       #instGetIoPart(ID := #hwID,   //read data from process image
                      OFFSET := #portAddr,
                      LEN := #statIOsize,
                      STATUS => #statIoPartStatus,
                      ERROR => #statIoPartError,
                      INPUTS := #statAnt);
       #statAntStatus := #statAnt[#INDEX_ANT_STATUS];    //status byte
       #statPresence := #statAntStatus.%X5;    //Presence bit. Transponder on field
   END_REGION

   REGION Check antenna status
       IF #statAnt[#INDEX_RFID_ERROR] <> 0 AND #statBusy THEN
           #tempStatus.%W0 := BYTE_TO_WORD(#statAnt[#INDEX_RFID_ERROR]);    //error_BLK
           #tempStatus.%W1 := #STATUS_ERROR_IDENT_RFID;                    //identifier rfid errors
           #statBusy := false;
           #tempDone := false;
           #tempError := TRUE;
           #statState := #STATE_IDLE;
       END_IF;
   END_REGION

   REGION Check execute
       REGION Idle
           IF NOT #execute THEN
               #tempDone := false;
               #tempError := false;
               #tempStatus := 0;
           END_IF;
       END_REGION

       REGION Job executed
           IF #execute AND #execute <> #statExecuteReq THEN //Positive Edge for antenna on
               #statBusy := TRUE;                              //Block active
               #tempDone := FALSE;                             //reset all output parameters
               #tempError := FALSE;
               #tempStatus := #STATUS_NO_JOB;
               IF #antennaState THEN                          //if antenna then activate the ANTENNA_ON process
                   #statState := #STATE_ANTENNA_ON;
               ELSIF NOT #antennaState THEN                   //if not antenna then activate the ANTENNA_OFF process 
                   #statState := #STATE_ANTENNA_OFF;
               END_IF;

           END_IF;
       END_REGION
       #statExecuteReq := #execute;
   END_REGION

   REGION State machine
       CASE #statState OF
           #STATE_IDLE:
               ;

           #STATE_ANTENNA_ON:  //Antenna_on
               //Antenna on process
               #statAntStatus.%X4 := false;                        //Reset Byte 0, bit 4
               #statSent[#INDEX_SEND_CMD] := #CMD_ANTENNA_ON;
               #instSetIoPart(ID := #hwID,                         //Write data into process image
                              OFFSET := #portAddr,
                              LEN := #statIOsize,
                              STATUS => #statIoPartStatus,
                              ERROR => #statIoPartError,
                              OUTPUTS := #statSent);
               IF NOT #statIoPartError AND #statAnt[#INDEX_RFID_ERROR] = 0 THEN
                   #statState := #STATE_READY;
               ELSIF #statIoPartError THEN
                   #tempError := true;
                   #statBusy := FALSE;
                   #tempStatus.%W0 := DWORD_TO_WORD(#statIoPartStatus);//error_BLK
                   #tempStatus.%W1 := #STATUS_ERROR_IDENT_BLOCK;                    //identifier block errors
                   #statState := #STATE_IDLE;
               END_IF;

           #STATE_ANTENNA_OFF:
               //Antenna off process
               #statAntStatus.%X4 := true;                         //set Byte 0, bit 4
               #statSent[#INDEX_SEND_CMD] := #CMD_ANTENNA_OFF;
               #instSetIoPart(ID := #hwID,                         //Write data into process image
                              OFFSET := #portAddr,
                              LEN := #statIOsize,
                              STATUS => #statIoPartStatus,
                              ERROR => #statIoPartError,
                              OUTPUTS := #statSent);
               IF NOT #statIoPartError AND #statAnt[#INDEX_RFID_ERROR] = 0 THEN
                   IF #statAntStatus = #CMD_ANTENNA_OFF THEN    //if status_byte=16#10 then antenna off
                       #statState := #STATE_READY;
                   END_IF;
               ELSIF #statIoPartError THEN
                   #tempError := true;
                   #statBusy := FALSE;
                   #tempStatus.%W0 := DWORD_TO_WORD(#statIoPartStatus);    //error_BLK
                   #tempStatus.%W1 := #STATUS_ERROR_IDENT_BLOCK;   //identifier block errors
                   #statState := #STATE_IDLE;
               END_IF;

           #STATE_READY:
               #tempDone := true;
               #statBusy := FALSE;
               #statState := #STATE_IDLE;
           ELSE
               #statState := #STATE_IDLE;
       END_CASE;
   END_REGION

   REGION Update output interface 
       #done := #tempDone;
       #busy := #statBusy;
       #error := #tempError;
       #status := #tempStatus;
       #presence := #statPresence;
   END_REGION
END_FUNCTION_BLOCK

FUNCTION_BLOCK "LIOLink_RF200_WriteTag"   // FB6, SCL
TITLE = LIOLink_RF200_WriteTag
{ S7_Optimized_Access := 'TRUE' }
AUTHOR : SIOS
FAMILY : LIOLink
VERSION : 2.4
// Writes tags on SIMATIC RF200 readers via IO-Link
   VAR_INPUT
      execute : Bool;   // Execute function
      addrTag : Word;   // Start address of data on tag
      length : Word;   // Length of data to be written
      hwID : HW_SUBMODULE;   // Hardware identifier of IO-Link communication module
      portAddr : Int;   // Start address of port
      "version" : USInt := 11;   // IO-Link version of the reader; 11: IO-Link V1.1, 10: IO-Link V1.0
   END_VAR
   VAR_OUTPUT
      done : Bool;   // TRUE: job done
      busy : Bool;   // FALSE: no job, TRUE: job in progress
      error : Bool;   // FALSE: no error, TRUE: error
      status : DWord;   // Error Status
      presence : Bool;   // Tag on antenna field
   END_VAR
   VAR_IN_OUT
      identData : Variant;   // Data to write in
   END_VAR
   VAR
      instTonR : TONR_TIME;   // Tag has left antenna field detection timer
      statState : Int;   // Main State Machine Index
      statTimerIn : Bool;   // Tag has left antenna field detection timer - Start Tag
      statTimerR : Bool;   // Tag has left antenna field detection timer - Reset Tag
      statTimerPt : Time := T#5S;   // Tag has left antenna field detection timer - Detection time
      statStatusByte : Byte;   // First received Byte from process image
      statDat : Array[0..#UPPER_BOUND_IO_FIELD] of Byte;   // Sent data
      statRecDat : Array[0..#UPPER_BOUND_IO_FIELD] of Byte;   // Received data
      statPresence : Bool;   // TRUE: Transponder on field
      statExecuteReq : Bool;   // State of execute input of last cycle
      statLength : DInt;   // Length of read Data
      statAddr : Word;   // Address of Tag
      statWriteOffset : Int;   // Data offset for write function
      statPresenceFf : Bool;   // Transpnder status of last cycle
      statWriteData : Array[0..#UPPER_BOUND_MAX_DATA_FIELD] of Byte;   // Data to write to tag
      statDiffToIOsizeNetto : Int;   // Difference to full IO size
      statBytemove : Int;   // Shift value for data
      statDone : Bool;   // TRUE: job done
      statBusy : Bool;   // FALSE: no job, TRUE: job in progress
      statError : Bool;   // FALSE: no error, TRUE: error
      instSetIoPart : SETIO_PART;   // Instance for PIQ writing
      statIoPartError : Bool;   // TRUE: data in process image is invalid
      statIoPartStatus : DWord;   // Status for IO access
      instGetIoPart : GETIO_PART;   // Instance for PII reading
      statReturnMoveBlkVar : Int;   // Return Value of Block Move
      statIOsize : USInt;   // Size of the IO-Link Master PII
      statIOsizeNetto : USInt;   // Size of the IO-Link Master PAE without header
   END_VAR
   VAR_TEMP
      tempStatus : DWord;   // Auxiliary tag for status output
   END_VAR
   VAR CONSTANT
      IOL_V10 : USInt := 10;   // Identifier IO-Link version 1.0
      IOL_V11 : USInt := 11;   // Identifier IO-Link version 1.1
      LEN_DATA_V10 : USInt := 8;   // Length of user data for IO-Link version 1.0
      LEN_DATA_V11 : USInt := 32;   // Length of user data for IO-Link version 1.1
      UPPER_BOUND_IO_FIELD : USInt := 31;   // Upper bound of Input and Output fields
      UPPER_BOUND_MAX_DATA_FIELD : UInt := 1999;   // Upper bound of the data field of a RFID Tag
      DATA_HEADER_SIZE : USInt := 4;   // IO-Link Header Size for version 1.0 and 1.1
      STATUS_ERROR_IDENT_BLOCK : Word := 16#0001;   // Error Identification for block internal faults
      STATUS_ERROR_IDENT_RFID : Word := 16#0011;   // Error Identification for RFID reader faults
      STATUS_NO_JOB : Word := 16#0000;   // No job requested
      STATUS_ERROR_TAG_HAS_LEFT : Word := 16#8101;   // Error - the RFID tag has left the reader
      STATUS_ERROR_STILL_ACTIVE : Word := 16#8102;   // Error - block still busy, no further request possible
      STATUS_ERROR_LENGTH : Word := 16#8104;   // Error - requested length is less than 0
      STATE_IDLE : Int := 0;   // State Machine - Idle State
      STATE_WRITE : Int := 2;   // State Machine - Read Tag
      STATE_TELEGRAM : Int := 1;   // State Machine - Prepare telegram
      STATE_ERROR : Int := 3;   // State Machine - Error State
      DETECTION_TIME_TAG_OFF_FIELD : Time := T#5S;   // Tag has left antenna field detection time
      CMD_WRITE : Byte := 16#01;   // Command to read data
      CMD_RESET : Byte := 16#00;   // Command to reset
      INDEX_CMD : USInt := 0;   // Index in DataField - Command
      INDEX_RFID_ERROR : USInt := 1;   // Index in DataField - Error
      INDEX_ADDR_HIGH : USInt := 2;   // Index in DataField - Address High Byte
      INDEX_ADDR_LOW : USInt := 3;   // Index in DataField - Address Low Byte
      INDEX_SOURCE_DATA : DInt := 4;   // Index in Data Field - Start of netto Data
      INDEX_REC_STATUS : DInt := 0;   // Index in Received DataField - Status
   END_VAR
   // statRecDat[0] := 16#0000;
   // statRecDat[1] := 16#0000;
   // statRecDat[2] := 16#00FF;
   // statRecDat[3] := 16#00FF;
BEGIN
   REGION BLOCK INFO HEADER
       //===============================================================================
       // Siemens / (c)Copyright 2022
       //-------------------------------------------------------------------------------
       // Title:            LIOLink_RF200_WriteTag
       // Function:         Writes tags on SIMATIC RF200 readers via IO-Link
       // Library:          LIOLink
       // Author:           Siemens Industry Online Support
       // Tested with:      CPU 1513-1 PN FW 2.8
       // Engineering:      TIA Portal V16
       // Restrictions:     --
       // Requirements:     --
       //-------------------------------------------------------------------------------
       // Change log table:
       // Version  | Date       | Expert in charge       | Changes applied
       //----------|------------|------------------------|------------------------------
       // 01.00.00 | 01.03.2015 | Online Support         | First release
       // 01.01.00 | 01.12.2016 | Online Support         | Upgrade to TIA Portal V14
       // 02.00.00 | 01.09.2017 | Online Support         | Upgrade to TIA Portal V14 SP1
       //                                                | Implementation of Programming styleguide
       //                                                | Added support for IO-Link V1.1 readers
       // 02.01.00 | 01.12.2017 | Online Support         | Bug fixes and performance improvements
       // 02.02.00 | 01.03.2020 | Online Support         | Upgrade to TIA Portal V16
       // 02.03.00 | 22.09.2020 | Online Support         | Integrated FB into LIOLink library
       //                                                | Renamed FB to LIOLink_RF200_WriteTag
       //                                                | Combined FBs for IO-Link V1.0 and V1.1
       //                                                | Minor bug fixes
       // 02.04.00 | 04.10.2022 | SUP SPH                | Optimization                                               
       //===============================================================================
   END_REGION

   REGION Check version
       IF #version = #IOL_V11 THEN   //determine IO-Link reader version (1.0/1.1) to set offsets
           #statIOsize := #LEN_DATA_V11;
           #statIOsizeNetto := #LEN_DATA_V11 - #DATA_HEADER_SIZE;
       ELSE
           #statIOsize := #LEN_DATA_V10;
           #statIOsizeNetto := #LEN_DATA_V10 - #DATA_HEADER_SIZE;
       END_IF;
   END_REGION

   REGION Get PII
       //read data from process image
       #instGetIoPart(ID := #hwID,
                      OFFSET := #portAddr,
                      LEN := #statIOsize,
                      STATUS => #statIoPartStatus,
                      ERROR => #statIoPartError,
                      INPUTS := #statRecDat);

       #statStatusByte := #statRecDat[#INDEX_REC_STATUS];    //Status Byte
       #statPresence := #statStatusByte.%X5;   //Presence bit. Transponder on field
   END_REGION

   REGION Check execute
       REGION Idle
           IF NOT #execute THEN
               #statDone := false;
               #statBusy := false;
               #statError := false;
               #tempStatus := #STATUS_NO_JOB;
           END_IF;
       END_REGION

       #statDiffToIOsizeNetto := WORD_TO_INT(#length) MOD #statIOsizeNetto;
       REGION Job requested
           IF #execute AND #execute <> #statExecuteReq THEN    //Positive edge for reading of data
               IF NOT #statBusy THEN
                   #statAddr := #addrTag;    //Transpoder Adress
                   #statLength := WORD_TO_DINT(#length);   //Length of read Data
                   #statState := #STATE_WRITE;
                   #statBusy := TRUE;
                   #statDone := FALSE;   //reset all the output parameters                                   
                   #statError := FALSE;
                   #tempStatus := #STATUS_NO_JOB;
                   #statWriteOffset := 0;
                   #statBytemove := 0;
                   //next step >> send write command
               ELSE
                   #tempStatus.%W0 := #STATUS_ERROR_STILL_ACTIVE;    //block is still active
                   #tempStatus.%W1 := #STATUS_ERROR_IDENT_BLOCK;   //Error identifier for block errors
                   #statState := #STATE_ERROR;
               END_IF;
               IF #length < USINT_TO_WORD(#statIOsizeNetto) THEN
                   #tempStatus.%W0 := #STATUS_ERROR_LENGTH;    //length too short
                   #tempStatus.%W1 := #STATUS_ERROR_IDENT_BLOCK;   //identifier rfid errors
                   #tempStatus := #tempStatus;
                   #statState := #STATE_ERROR;
               END_IF;
           END_IF;
       END_REGION
       #statExecuteReq := #execute;
   END_REGION

   REGION Tag presence detection
       IF NOT #statPresence AND #statPresence <> #statPresenceFf THEN    //the tag has left the antenna  field
           IF NOT #statDone THEN
               #statTimerIn := true;   //wait 5 sec
               #statTimerR := false;
           END_IF;
       END_IF;
       #statPresenceFf := #statPresence;
       IF #statPresence THEN
           #statTimerR := true;
           #statTimerIn := false;
       END_IF;
   END_REGION

   REGION State machine
       CASE #statState OF
           #STATE_IDLE:
               #statWriteOffset := 0;    //offset of puffer must be reseted
               #statBusy := false;
               #statTimerIn := false;

           #STATE_WRITE:
               IF #statLength > 0 THEN
                   #statDat[#INDEX_CMD] := #CMD_WRITE;   //Set write command
                   #statDat[#INDEX_ADDR_HIGH] := #statAddr.%B1;    //Adr-H
                   #statDat[#INDEX_ADDR_LOW] := #statAddr.%B0;   //Adr-L
                   VariantGet(SRC := #identData,
                              DST => #statWriteData);

                   #statReturnMoveBlkVar := MOVE_BLK_VARIANT(SRC := #statWriteData,
                                                             COUNT := #statIOsizeNetto,
                                                             SRC_INDEX := #statWriteOffset - #statBytemove,
                                                             DEST_INDEX := #INDEX_SOURCE_DATA,
                                                             DEST => #statDat);
                   //Just #statIOsizeNetto Bytes are reserved for every transfer
               END_IF;
               IF NOT #statIoPartError THEN
                   #statState := #STATE_TELEGRAM;    //Telegram: Edit the read data
               END_IF;

           #STATE_TELEGRAM:
               IF #statLength > 0 THEN   //Only when length of data>0 can continue  
                   IF #statStatusByte.%X6 THEN   //IF RFID error has occured
                       #tempStatus.%W0 := #statRecDat[#INDEX_RFID_ERROR];
                       #tempStatus.%W1 := #STATUS_ERROR_IDENT_RFID;    //Error identifier for RFID errors
                       #statState := #STATE_ERROR;
                   END_IF;

                   //-------------------------- write command is ready------------------------------------------------//
                   IF #statStatusByte.%X7 AND #statStatusByte.%X0 THEN
                       IF #statRecDat[#INDEX_ADDR_HIGH] = #statAddr.%B1 AND #statRecDat[#INDEX_ADDR_LOW] = #statAddr.%B0 THEN //received ADR must be ==sent ADR

                           IF NOT #statIoPartError THEN
                               IF #statStatusByte.%X7 AND NOT #statStatusByte.%X6 THEN
                                   #statLength := #statLength - #statIOsizeNetto;
                                   IF #statDiffToIOsizeNetto <> 0 AND #statLength < #statIOsizeNetto THEN
                                       #statBytemove := #statIOsizeNetto - #statDiffToIOsizeNetto;
                                   END_IF;
                                   //if len is not dividable with #statIOsizeNetto the adr offset has to be changed that the last (length < #statIOsizeNetto) command is done right
                                   #statWriteOffset := #statWriteOffset + #statIOsizeNetto;                                   //offset must be changed
                                   #statAddr := INT_TO_WORD(WORD_TO_INT(#statAddr) + USINT_TO_INT(#statIOsizeNetto) - #statBytemove);     //Change the ADR on Transponder(#statIOsizeNetto Bytes)       
                                   #statState := #STATE_WRITE;                      //Start a new write command
                               ELSE
                                   #statState := #STATE_IDLE;
                               END_IF;
                           ELSE
                               #tempStatus.%W0 := DWORD_TO_WORD(#statIoPartStatus);    //Error has to BLKMOV occured
                               #tempStatus.%W1 := #STATUS_ERROR_IDENT_BLOCK;   //functions-Error identifier
                               #statState := #STATE_ERROR;
                           END_IF;
                       END_IF;
                   END_IF;

                   #instSetIoPart(ID := #hwID,
                                  OFFSET := #portAddr,
                                  LEN := #statIOsize,
                                  STATUS => #statIoPartStatus,
                                  ERROR => #statIoPartError,
                                  OUTPUTS := #statDat);

                   IF #statIoPartError THEN
                       #tempStatus.%W0 := DWORD_TO_WORD(#statIoPartStatus);   //Error has to BLKMOV occured
                       #tempStatus.%W1 := #STATUS_ERROR_IDENT_BLOCK;   //functions-Error identifier
                       #statState := #STATE_ERROR;
                   END_IF;

               ELSE
                   #statState := #STATE_IDLE;
                   #statBusy := false;
                   #statDone := TRUE;

                   //Reset write command
                   #statDat[#INDEX_CMD] := #CMD_RESET;

                   #instSetIoPart(ID := #hwID,
                                  OFFSET := #portAddr,
                                  LEN := #statIOsize,
                                  STATUS => #statIoPartStatus,
                                  ERROR => #statIoPartError,
                                  OUTPUTS := #statDat);
               END_IF;

           #STATE_ERROR:
               #statError := TRUE;
               #statBusy := false;
               #statDone := false;
               #statTimerIn := false;
               #statTimerR := true;
               #statState := #STATE_IDLE;

               //Reset write command
               #statDat[#INDEX_CMD] := #CMD_RESET;

               #instSetIoPart(ID := #hwID,
                              OFFSET := #portAddr,
                              LEN := #statIOsize,
                              STATUS => #statIoPartStatus,
                              ERROR => #statIoPartError,
                              OUTPUTS := #statDat);
           ELSE
               #statState := #STATE_IDLE;
       END_CASE;
   END_REGION

   REGION Detection timer
       #instTonR(IN := #statTimerIn,   //this timer will start, if the tag has left the antenna field
                 R := #statTimerR,
                 PT := #statTimerPt);
       IF #instTonR.Q THEN   //error has occured. No tag on field during the 5 sec.
           #tempStatus.%W0 := #STATUS_ERROR_TAG_HAS_LEFT;  //tag has left the field
           #tempStatus.%W1 := #STATUS_ERROR_IDENT_BLOCK;   //identifier rfid errors
           #statState := #STATE_ERROR;
       END_IF;
   END_REGION

   REGION Update output interface 
       #done := #statDone;
       #busy := #statBusy;
       #error := #statError;
       #status := #tempStatus;
       #presence := #statPresence;
   END_REGION
END_FUNCTION_BLOCK

FUNCTION_BLOCK "LIOLink_RF200"   // FB5200, SCL
TITLE = LIOLink_RF200 / IO_LINK_RFID_1500
{ S7_Optimized_Access := 'TRUE' }
AUTHOR : SIOS
FAMILY : LIOLink
VERSION : 3.0
// IO-Link Device FB for SIMATIC RF200 to use with S7-1200/1500 controllers! / IO-Link Geraete FB fuer SIMATIC RFID zur Nutzung mit S7-1500!
   VAR_INPUT
      execute : Bool;   // Request job (on rising edge)
      hwID : HW_IO;   // Hardware identifier of IO-Link master module or first sub module
      cap : Int;   // Client Access Point (CAP) 0xB400 or 0x00E3 (227)
      readWrite : Bool;   // Read and write access to IO-Link device 0: Read, 1:Write
      port : Int;   // Port of device on the IO-Link Master
      pollingPeriod : Time := T#100MS;   // Time period of polling
      directParameter1 : Bool;   // Read parameter page 1
      systemCommand : Bool;   // Read system commands
      deviceAccessLocks : Bool;   // Read device access locks
      vendorName : Bool;   // Read manufacturer name
      vendorText : Bool;   // Read manufacturer text
      productName : Bool;   // Read product name
      productID : Bool;   // Read product ID
      productText : Bool;   // Read product text
      serialNumber : Bool;   // Read serial number
      hwRevision : Bool;   // Read hardware revision
      fwRevision : Bool;   // Read firmware revision
      appSpecificName : Bool;   // Read/Write application specific name
      errorCount : Bool;   // Read error count
      deviceStatus : Bool;   // Read device status
      deviceStatusDetailed : Bool;   // Read device status detailed
      processIn : Bool;   // Read process data IN
      processOut : Bool;   // Read process data OUT
      parameters : Bool;   // Read parameters
      eventHistory : Bool;   // Read event history
      readerStatus : Bool;   // Read status of reader
      tagStatus : Bool;   // Reag tag status
      uidHistory : Bool;   // Read UID history
   END_VAR
   VAR_OUTPUT
      done : Bool;   // 0: data invalid, 1: data valid
      busy : Bool;   // 0: job done, 1: job in progress
      error : Bool;   // 0: no error, 1: error
      status : Word;   // DP/PN IO error status
      diagnostics : "LIOLink_typeDiagnostics";   // IO-Link error status
   END_VAR
   VAR_IN_OUT
      data : "LIOLink_RF200_typeAll";   // Device data buffer
   END_VAR
   VAR
      instDevice : "LIOLink_Device";
      statRecordParam : Struct   // Data set parameters
         index : Array[0..#HIGHEST_REQUEST_NUMBER] of Int;   // Data set index
         subindex : Array[0..#HIGHEST_REQUEST_NUMBER] of Int;   // Data set subindex
         length : Array[0..#HIGHEST_REQUEST_NUMBER] of Int;   // Data set length
      END_STRUCT;
      statRecord : Array[0..#UPPER_BOUND_RECORD] of Byte;   // Record buffer
      statIndex : Int;   // Requested index
      statSubindex : Int;   // Requested subindex
      statRecordLen : Int;   // Length of record to be written
      statHwID : HW_IO;   // Static value for input 'hwID'
      statCap : Int;   // Static value for input 'cap'
      statReadWrite : Bool;   // Static value for input 'readWrite'
      statPort : Int;   // Static value for input 'port'
      statPollingPeriod : Time;   // Static value for input 'pollingPeriod'
      statDirectParameter1 : Bool;   // Static value for input 'directParameter1'
      statSystemCommand : Bool;   // Static value for input 'systemCommands'
      statDeviceAccessLocks : Bool;   // Static value for input 'deviceAccessLocks'
      statVendorName : Bool;   // Static value for input 'vendorName'
      statVendorText : Bool;   // Static value for input 'vendorText'
      statProductName : Bool;   // Static value for input 'productName'
      statProductID : Bool;   // Static value for input 'productID'
      statProductText : Bool;   // Static value for input 'productText'
      statSerialNumber : Bool;   // Static value for input 'serialNumber'
      statHwRevision : Bool;   // Static value for input 'hwRevision'
      statFwRevision : Bool;   // Static value for input 'fwRevision'
      statAppSpecificName : Bool;   // Static value for input 'appSpecificName'
      statErrorCount : Bool;   // Static value for input 'errorCount'
      statDeviceStatus : Bool;   // Static value for input 'deviceStatus'
      statDeviceStatusDetailed : Bool;   // Static value for input 'deviceStatusDetailed'
      statProcessIn : Bool;   // Static value for input 'processIn'
      statProcessOut : Bool;   // Static value for input 'processOut'
      statParameters : Bool;   // Static value for input 'parameters'
      statEventHistory : Bool;   // Static value for input 'eventHistory'
      statReaderStatus : Bool;   // Static value for input 'readerStatus'
      statTagStatus : Bool;   // Static value for input 'tagStatus'
      statUidHistory : Bool;   // Static value for input 'uidHistory'
      statRequest : Int;   // Case of request (data set)
      statDoneOld : Bool;   // Last cycle's value of instDevice.done
   END_VAR
   VAR_TEMP
      tempIndex : UInt;   // Loop index
      tempLen : UInt;   // Auxiliary tag Length
      tempRetValSerialize : Int;   // Auxiliary tag for Serialize RetVal
      tempRetValDeserialize : Int;   // Auxiliary tag for Deserialize RetVal
      tempPosSerialize : DInt;   // Auxiliary tag for Serialize POS
      tempPosDeserialize : DInt;   // Auxiliary tag for Deserialize POS Output
      tempFieldParameterPage0 : Array[0..#UPPER_BOUND_PARAMETER_PAGE0] of Byte;   // Auxiliary tag for Parameter Page 0 record conversion
      tempFieldParameters : Array[0..#UPPER_BOUND_PARAMETERS] of Byte;   // Auxiliary tag for Parameters record conversion
      tempFieldEventHistory : Array[0..#UPPER_BOUND_EVENT_HISTORY] of Byte;   // Auxiliary tag for EventHistory record conversion
      tempFieldReaderStatus : Array[0..#UPPER_BOUND_READER_STATUS] of Byte;   // Auxiliary tag for Reader Status record conversion
      tempFieldTagStatus : Array[0..#UPPER_BOUND_TAG_STATUS] of Byte;   // Auxiliary tag for Tag Status record conversion
      tempFieldUIDHistory : Array[0..#UPPER_BOUND_UID_HISTORY] of Byte;   // Auxiliary tag for UID History record conversion
      tempInternalError : Bool;   // Auxiliary tag to collect serialize and Deserialize issues
   END_VAR
   VAR CONSTANT
      UPPER_BOUND_RECORD : Int := 231;   // Upper Bound of record buffer
      HIGHEST_REQUEST_NUMBER : Int := 28;   // Highest available request number
      UPPER_BOUND_PARAMETER_PAGE0 : Int := 15;   // Upper Bound of Parameter Page 0 auxiliary field
      UPPER_BOUND_PARAMETERS : Int := 7;   // Upper Bound of Parameters auxiliary field
      UPPER_BOUND_EVENT_HISTORY : Int := 19;   // Upper Bound of Event History auxiliary field
      UPPER_BOUND_READER_STATUS : Int := 17;   // Upper Bound of Reader Status auxiliary field
      UPPER_BOUND_TAG_STATUS : Int := 15;   // Upper Bound of Tag Status auxiliary field
      UPPER_BOUND_UID_HISTORY : Int := 39;   // Upper Bound of UID History auxiliary field
      MODE_READ : Bool := FALSE;   // Mode to read data
      MODE_WRITE : Bool := TRUE;   // Mode to write data
      STATUS_IDLE : Word := 16#7000;   // Status: Idle
      STATUS_EXECUTION_FINISHED : Word := 16#0000;   // Execution finished without errors
      ERR_INCONSISTENT_DATA : Word := 16#8402;   // Error: Read data record doesn't match request
      INDEX_DIRECT_PARAM1 : Int := 0;   // Record Index
      INDEX_SYSTEM_COMMAND : Int := 2;   // Record Index
      INDEX_ACCESS_LOCKS : Int := 12;   // Record Index
      INDEX_EVENT_HISTORY : Int := 74;   // Record Index
      INDEX_VENDOR_NAME : Int := 16;   // Record Index
      INDEX_VENDOR_TEXT : Int := 17;   // Record Index
      INDEX_PRODUCT_NAME : Int := 18;   // Record Index
      INDEX_PRODUCT_ID : Int := 19;   // Record Index
      INDEX_PRODUCT_TEXT : Int := 20;   // Record Index
      INDEX_SERIAL_NUMBER : Int := 21;   // Record Index
      INDEX_HARDWARE_REVISION : Int := 22;   // Record Index
      INDEX_FIRMWARE_REVISION : Int := 23;   // Record Index
      INDEX_APP_SPECIFIC_NAME : Int := 24;   // Record Index
      INDEX_ERROR_COUNT : Int := 32;   // Record Index
      INDEX_DEVICE_STATUS : Int := 36;   // Record Index
      INDEX_DETAILED_STATUS : Int := 37;   // Record Index
      INDEX_PII : Int := 40;   // Record Index
      INDEX_PIQ : Int := 41;   // Record Index
      INDEX_PARAMETERS : Int := 64;   // Record Index
      INDEX_TAG_STATUS : Int := 91;   // Record Index
      INDEX_READER_STATUS : Int := 90;   // Record Index
      INDEX_UID_HISTORY : Int := 92;   // Record Index
      LENGTH_DIRECT_PARAM1 : Int := 16;   // Record Length
      LENGTH_SYSTEM_COMMAND : Int := 1;   // Record Length
      LENGTH_ACCESS_LOCKS : Int := 2;   // Record Length
      LENGTH_EVENT_HISTORY : Int := 20;   // Record Length
      LENGTH_VENDOR_NAME : Int := 12;   // Record Length
      LENGTH_VENDOR_TEXT : Int := 12;   // Record Length
      LENGTH_PRODUCT_NAME : Int := 24;   // Record Length
      LENGTH_PRODUCT_ID : Int := 16;   // Record Length
      LENGTH_PRODUCT_TEXT : Int := 64;   // Record Length
      LENGTH_SERIAL_NUMBER : Int := 12;   // Record Length
      LENGTH_HARDWARE_REVISION : Int := 12;   // Record Length
      LENGTH_FIRMWARE_REVISION : Int := 12;   // Record Length
      LENGTH_APP_SPECIFIC_NAME : Int := 32;   // Record Length
      LENGTH_ERROR_COUNT : Int := 2;   // Record Length
      LENGTH_DEVICE_STATUS : Int := 1;   // Record Length
      LENGTH_DETAILED_STATUS : Int := 1;   // Record Length
      LENGTH_PII : Int := 8;   // Record Length
      LENGTH_PIQ : Int := 8;   // Record Length
      LENGTH_PARAMETERS : Int := 8;   // Record Length
      LENGTH_TAG_STATUS : Int := 15;   // Record Length
      LENGTH_READER_STATUS : Int := 18;   // Record Length
      LENGTH_UID_HISTORY : Int := 40;   // Record Length
      EMPTY_CHAR : Char := '$00';   // Default empty chat to fill empty field entries
      DEVICE_TIMEOUT : Time := T#20S;   // Timeout value for the IO-Link Device Instance
   END_VAR
   // statRecordParam.index[0] := 0;
   // statRecordParam.index[1] := 0;
   // statRecordParam.index[2] := 0;
   // statRecordParam.index[3] := 0;
   // statRecordParam.index[4] := 0;
   // statRecordParam.index[5] := 0;
   // statRecordParam.index[6] := 0;
   // statRecordParam.index[7] := 0;
   // statRecordParam.index[8] := 0;
   // statRecordParam.index[9] := 74;
   // statRecordParam.index[10] := 16;
   // statRecordParam.index[11] := 17;
   // statRecordParam.index[12] := 18;
   // statRecordParam.index[13] := 19;
   // statRecordParam.index[14] := 20;
   // statRecordParam.index[15] := 21;
   // statRecordParam.index[16] := 22;
   // statRecordParam.index[17] := 23;
   // statRecordParam.index[18] := 24;
   // statRecordParam.index[19] := 32;
   // statRecordParam.index[20] := 0;
   // statRecordParam.index[21] := 0;
   // statRecordParam.index[22] := 91;
   // statRecordParam.index[23] := 90;
   // statRecordParam.index[24] := 92;
   // statRecordParam.index[25] := 0;
   // statRecordParam.index[26] := 0;
   // statRecordParam.index[27] := 0;
   // statRecordParam.index[28] := 0;
   // statRecordParam.length[0] := 0;
   // statRecordParam.length[1] := 16;
   // statRecordParam.length[2] := 0;
   // statRecordParam.length[3] := 0;
   // statRecordParam.length[4] := 0;
   // statRecordParam.length[5] := 0;
   // statRecordParam.length[6] := 0;
   // statRecordParam.length[7] := 0;
   // statRecordParam.length[8] := 0;
   // statRecordParam.length[9] := 20;
   // statRecordParam.length[10] := 12;
   // statRecordParam.length[11] := 12;
   // statRecordParam.length[12] := 24;
   // statRecordParam.length[13] := 16;
   // statRecordParam.length[14] := 0;
   // statRecordParam.length[15] := 0;
   // statRecordParam.length[16] := 0;
   // statRecordParam.length[17] := 12;
   // statRecordParam.length[18] := 32;
   // statRecordParam.length[19] := 2;
   // statRecordParam.length[20] := 0;
   // statRecordParam.length[21] := 0;
   // statRecordParam.length[22] := 15;
   // statRecordParam.length[23] := 18;
   // statRecordParam.length[24] := 40;
   // statRecordParam.length[25] := 0;
   // statRecordParam.length[26] := 0;
   // statRecordParam.length[27] := 0;
   // statRecordParam.length[28] := 0;
BEGIN
   REGION BLOCK INFO HEADER
       //===============================================================================
       // Siemens / (c)Copyright 2023
       //-------------------------------------------------------------------------------
       // Title:            LIOLink_RF200
       // Function:         Capsule block to communicate with SIMATIC RF200 Readers
       // Library:          LIOLink
       // Author:           Siemens Industry Online Support
       // Tested with:      CPU 1513-1 PN FW 2.8
       // Engineering:      TIA Portal V16
       // Restrictions:     --
       // Requirements:     --
       //-------------------------------------------------------------------------------
       // Change log table:
       // Version  | Date       | Expert in charge       | Changes applied
       //----------|------------|------------------------|------------------------------
       // 01.00.00 | 11.04.2014 | Online Support         | First release
       // 02.00.00 | 30.03.2015 | Online Support         | Upgrade to TIA Portal V13 SP1, use function IO_LINK_DEVICE, only one function for S7-1200 and 1500
       // 02.01.00 | 23.10.2015 | Online Support         | Update to IO_LINK_DEVICE Version 3.1
       // 03.00.00 | 01.09.2020 | Online Support         | Rewrote block for FB "LIOLink_Device" V4.0.0
       // 03.01.00 | 25.10.2022 | SUP SPH                | Optimized and function extension
       //===============================================================================
   END_REGION

   REGION INIT
       IF (#execute = TRUE AND #instDevice.status = #STATUS_IDLE) THEN

           REGION Inputs
               //save inputs
               #statHwID := #hwID;
               #statCap := #cap;
               #statReadWrite := #readWrite;
               #statPort := #port;
               #statPollingPeriod := #pollingPeriod;
               #statDirectParameter1 := #directParameter1;
               #statSystemCommand := #systemCommand;
               #statDeviceAccessLocks := #deviceAccessLocks;
               #statVendorName := #vendorName;
               #statVendorText := #vendorText;
               #statProductName := #productName;
               #statProductID := #productID;
               #statProductText := #productText;
               #statSerialNumber := #serialNumber;
               #statHwRevision := #hwRevision;
               #statFwRevision := #fwRevision;
               #statAppSpecificName := #appSpecificName;
               #statErrorCount := #errorCount;
               #statDeviceStatus := #deviceStatus;
               #statDeviceStatusDetailed := #deviceStatusDetailed;
               #statProcessIn := #processIn;
               #statProcessOut := #processOut;
               #statParameters := #parameters;
               #statEventHistory := #eventHistory;
               #statReaderStatus := #readerStatus;
               #statTagStatus := #tagStatus;
               #statUidHistory := #uidHistory;
           END_REGION

           REGION Request selector
               //set Index and RecordLen based on the request
               IF #statDirectParameter1 THEN
                   #statIndex := #INDEX_DIRECT_PARAM1;
                   #statRecordLen := #LENGTH_DIRECT_PARAM1;
               ELSIF #statSystemCommand THEN
                   #statIndex := #INDEX_SYSTEM_COMMAND;
                   #statRecordLen := #LENGTH_SYSTEM_COMMAND;
               ELSIF #statDeviceAccessLocks THEN
                   #statIndex := #INDEX_ACCESS_LOCKS;
                   #statRecordLen := #LENGTH_ACCESS_LOCKS;
               ELSIF #statVendorName THEN
                   #statIndex := #INDEX_VENDOR_NAME;
                   #statRecordLen := #LENGTH_VENDOR_NAME;
               ELSIF #statVendorText THEN
                   #statIndex := #INDEX_VENDOR_TEXT;
                   #statRecordLen := #LENGTH_VENDOR_TEXT;
               ELSIF #statProductName THEN
                   #statIndex := #INDEX_PRODUCT_NAME;
                   #statRecordLen := #LENGTH_PRODUCT_NAME;
               ELSIF #statProductID THEN
                   #statIndex := #INDEX_PRODUCT_ID;
                   #statRecordLen := #LENGTH_PRODUCT_ID;
               ELSIF #statProductText THEN
                   #statIndex := #INDEX_PRODUCT_TEXT;
                   #statRecordLen := #LENGTH_PRODUCT_TEXT;
               ELSIF #statSerialNumber THEN
                   #statIndex := #INDEX_SERIAL_NUMBER;
                   #statRecordLen := #LENGTH_SERIAL_NUMBER;
               ELSIF #statHwRevision THEN
                   #statIndex := #INDEX_HARDWARE_REVISION;
                   #statRecordLen := #LENGTH_HARDWARE_REVISION;
               ELSIF #statFwRevision THEN
                   #statIndex := #INDEX_FIRMWARE_REVISION;
                   #statRecordLen := #LENGTH_FIRMWARE_REVISION;
               ELSIF #statAppSpecificName THEN
                   #statIndex := #INDEX_APP_SPECIFIC_NAME;
                   #statRecordLen := #LENGTH_APP_SPECIFIC_NAME;
               ELSIF #statErrorCount THEN
                   #statIndex := #INDEX_ERROR_COUNT;
                   #statRecordLen := #LENGTH_ERROR_COUNT;
               ELSIF #statDeviceStatus THEN
                   #statIndex := #INDEX_DEVICE_STATUS;
                   #statRecordLen := #LENGTH_DEVICE_STATUS;
               ELSIF #statDeviceStatusDetailed THEN
                   #statIndex := #INDEX_DETAILED_STATUS;
                   #statRecordLen := #LENGTH_DETAILED_STATUS;
               ELSIF #statProcessIn THEN
                   #statIndex := #INDEX_PII;
                   #statRecordLen := #LENGTH_PII;
               ELSIF #statProcessOut THEN
                   #statIndex := #INDEX_PIQ;
                   #statRecordLen := #LENGTH_PIQ;
               ELSIF #statParameters THEN
                   #statIndex := #INDEX_PARAMETERS;
                   #statRecordLen := #LENGTH_PARAMETERS;
               ELSIF #statEventHistory THEN
                   #statIndex := #INDEX_EVENT_HISTORY;
                   #statRecordLen := #LENGTH_EVENT_HISTORY;
               ELSIF #statReaderStatus THEN
                   #statIndex := #INDEX_READER_STATUS;
                   #statRecordLen := #LENGTH_READER_STATUS;
               ELSIF #statTagStatus THEN
                   #statIndex := #INDEX_TAG_STATUS;
                   #statRecordLen := #LENGTH_TAG_STATUS;
               ELSIF #statUidHistory THEN
                   #statIndex := #INDEX_UID_HISTORY;
                   #statRecordLen := #LENGTH_UID_HISTORY;
               ELSE
                   RETURN;
               END_IF;
           END_REGION

           IF #statReadWrite = #MODE_WRITE THEN
               //prepare statRecord in case of a writing request
               REGION write
                   IF #statSystemCommand THEN
                       #statRecord[0] := #data.systemCommand;

                   ELSIF #statDeviceAccessLocks THEN
                       #statRecord[0] := #data.deviceAccessLocks.%B0;
                       #statRecord[1] := #data.deviceAccessLocks.%B1;

                   ELSIF #statAppSpecificName THEN
                       Strg_TO_Chars(Strg := #data.appSpecificName,
                                     pChars := 0,
                                     Cnt => #tempLen,
                                     Chars := #statRecord);

                   ELSIF #statParameters THEN
                       #tempRetValSerialize := Serialize(SRC_VARIABLE := #data.parameters, DEST_ARRAY => #tempFieldParameters, POS := #tempPosSerialize);
                       UMOVE_BLK(IN := #tempFieldParameters[0],
                                 COUNT := INT_TO_ULINT(#statRecordLen),
                                 OUT => #statRecord[0]);
                       // Fill remaining characters with null
                       FOR #tempIndex := #tempLen TO INT_TO_UINT(#statRecordLen - 1) DO
                           #statRecord[#tempIndex] := CHAR_TO_BYTE(#EMPTY_CHAR);
                       END_FOR;
                   ELSE // all other data sets are read only  
                       ;
                   END_IF;
                   #tempInternalError := #tempRetValSerialize <> WORD_TO_INT(#STATUS_EXECUTION_FINISHED);
               END_REGION
           END_IF;
       END_IF;
   END_REGION

   REGION CALL
       //IOL-Call -> Request to read/write from an IO-Link-Device
       #instDevice(execute := #execute,
                   hwID := #statHwID,
                   cap := #statCap,
                   readWrite := #statReadWrite,
                   "port" := #statPort,
                   pollingPeriod := #statPollingPeriod,
                   index := #statIndex,
                   subindex := #statSubindex,
                   writeLen := #statRecordLen,
                   timeout := #DEVICE_TIMEOUT,
                   record := #statRecord);
   END_REGION

   REGION READ
       // Copy data if available and valid
       IF #instDevice.done = TRUE AND #statDoneOld = FALSE AND #statReadWrite = #MODE_READ THEN
           IF #statDirectParameter1 THEN
               UMOVE_BLK(IN := #statRecord[0],
                         COUNT := INT_TO_ULINT(#statRecordLen),
                         OUT => #tempFieldParameterPage0[0]);
               #tempRetValDeserialize := Deserialize(SRC_ARRAY := #tempFieldParameterPage0, DEST_VARIABLE => #data.directParameterPage, POS := #tempPosDeserialize);

           ELSIF #statDeviceAccessLocks THEN
               #data.deviceAccessLocks.%B0 := #statRecord[0];
               #data.deviceAccessLocks.%B1 := #statRecord[1];

           ELSIF #statVendorName THEN
               Chars_TO_Strg(Chars := #statRecord,
                             pChars := 0,
                             Cnt := INT_TO_UINT(#statRecordLen),
                             Strg => #data.vendorName);

           ELSIF #statVendorText THEN
               Chars_TO_Strg(Chars := #statRecord,
                             pChars := 0,
                             Cnt := INT_TO_UINT(#statRecordLen),
                             Strg => #data.vendorText);

           ELSIF #statProductName THEN
               Chars_TO_Strg(Chars := #statRecord,
                             pChars := 0,
                             Cnt := INT_TO_UINT(#statRecordLen),
                             Strg => #data.productName);

           ELSIF #statProductID THEN
               Chars_TO_Strg(Chars := #statRecord,
                             pChars := 0,
                             Cnt := INT_TO_UINT(#statRecordLen),
                             Strg => #data.productID);

           ELSIF #statProductText THEN
               Chars_TO_Strg(Chars := #statRecord,
                             pChars := 0,
                             Cnt := INT_TO_UINT(#statRecordLen),
                             Strg => #data.productText);

           ELSIF #statSerialNumber THEN
               Chars_TO_Strg(Chars := #statRecord,
                             pChars := 0,
                             Cnt := INT_TO_UINT(#statRecordLen),
                             Strg => #data.serialNumber);

           ELSIF #statHwRevision THEN
               Chars_TO_Strg(Chars := #statRecord,
                             pChars := 0,
                             Cnt := INT_TO_UINT(#statRecordLen),
                             Strg => #data.hwRevision);

           ELSIF #statFwRevision THEN
               Chars_TO_Strg(Chars := #statRecord,
                             pChars := 0,
                             Cnt := INT_TO_UINT(#statRecordLen),
                             Strg => #data.fwRevision);

           ELSIF #statAppSpecificName THEN
               Chars_TO_Strg(Chars := #statRecord,
                             pChars := 0,
                             Cnt := INT_TO_UINT(#statRecordLen),
                             Strg => #data.appSpecificName);

           ELSIF #statErrorCount THEN
               #data.errorCount.%B0 := #statRecord[1];
               #data.errorCount.%B1 := #statRecord[0];

           ELSIF #statDeviceStatus THEN
               #data.deviceStatus := #statRecord[0];

           ELSIF #statDeviceStatusDetailed THEN
               #data.deviceStatusDetailed := #statRecord[0];

           ELSIF #statProcessIn THEN
               UMOVE_BLK(IN := #statRecord[0],
                         COUNT := INT_TO_ULINT(#statRecordLen),
                         OUT => #data.processImageIn[0]);

           ELSIF #statProcessOut THEN
               UMOVE_BLK(IN := #statRecord[0],
                         COUNT := INT_TO_ULINT(#statRecordLen),
                         OUT => #data.processImageOut[0]);

           ELSIF #statParameters THEN
               UMOVE_BLK(IN := #statRecord[0],
                         COUNT := INT_TO_ULINT(#statRecordLen),
                         OUT => #tempFieldParameters[0]);
               #tempRetValDeserialize := Deserialize(SRC_ARRAY := #tempFieldParameters, DEST_VARIABLE => #data.parameters, POS := #tempPosDeserialize);

           ELSIF #statEventHistory THEN
               UMOVE_BLK(IN := #statRecord[0],
                         COUNT := INT_TO_ULINT(#statRecordLen),
                         OUT => #tempFieldEventHistory[0]);
               #tempRetValDeserialize := Deserialize(SRC_ARRAY := #tempFieldEventHistory, DEST_VARIABLE => #data.eventHistory, POS := #tempPosDeserialize);

           ELSIF #statReaderStatus THEN
               UMOVE_BLK(IN := #statRecord[0],
                         COUNT := INT_TO_ULINT(#statRecordLen),
                         OUT => #tempFieldReaderStatus[0]);
               #tempRetValDeserialize := Deserialize(SRC_ARRAY := #tempFieldReaderStatus, DEST_VARIABLE => #data.readerStatus, POS := #tempPosDeserialize);

           ELSIF #statTagStatus THEN
               UMOVE_BLK(IN := #statRecord[0],
                         COUNT := INT_TO_ULINT(#statRecordLen),
                         OUT => #tempFieldTagStatus[0]);
               #tempRetValDeserialize := Deserialize(SRC_ARRAY := #tempFieldTagStatus, DEST_VARIABLE => #data.tagStatus, POS := #tempPosDeserialize);

           ELSIF #statUidHistory THEN
               UMOVE_BLK(IN := #statRecord[0],
                         COUNT := INT_TO_ULINT(#statRecordLen),
                         OUT => #tempFieldUIDHistory[0]);
               #tempRetValDeserialize := Deserialize(SRC_ARRAY := #tempFieldUIDHistory, DEST_VARIABLE => #data.uidHistory, POS := #tempPosDeserialize);
           ELSE // Other data sets are not defined
               ;
           END_IF;
           #tempInternalError := #tempRetValDeserialize <> WORD_TO_INT(#STATUS_EXECUTION_FINISHED);
       END_IF;

       #statDoneOld := #instDevice.done;
   END_REGION

   REGION OUTPUTS
       IF #tempInternalError THEN //Error occured
           #done := false;
           #busy := false;
           #error := true;
           #status := #ERR_INCONSISTENT_DATA;
       ELSE //Execute successful
           #done := #instDevice.done;
           #busy := #instDevice.busy;
           #error := #instDevice.error;
           #status := #instDevice.status;
           #diagnostics := #instDevice.diagnostics;
       END_IF;
   END_REGION
END_FUNCTION_BLOCK

// folder: LIOLink/S7-1200/1500/Device-specific blocks/SIRIUS

FUNCTION_BLOCK "LIOLink_3RA"   // FB5100, SCL
TITLE = LIOLink_3RA / IO_LINK_3RAxy
{ S7_Optimized_Access := 'TRUE' }
AUTHOR : SIOS
FAMILY : LIOLink
VERSION : 3.1
// IO-Link Device FB for SIRIUS 3RAxy to use with S7-1200/1500 controllers! / IO-Link Geraete FB fuer SIRIUS 3RAxy zur Nutzung mit S7-1500!
   VAR_INPUT
      execute : Bool;   // Request to execute function
      cap : Int;   // Client Access Point (CAP) 0xB400 or 0x00E3 (227)
      hwID : HW_IO;   // Hardware identifier of IO-Link master module or first sub module
      readWrite : Bool;   // FALSE: read, TRUE: write
      port : Int;   // Port of the IO-Link Master for the Device
      pollingPeriod : Time := T#100MS;   // Time period of polling
      parameterPage0 : Bool;   // Read access on parameter page 0
      parameterPage1 : Bool;   // Read/Write access on parameter page 1
      vendorName : Bool;   // Read Vendor Name
      vendorText : Bool;   // Read Vendor Text
      productName : Bool;   // Read Product Name
      productID : Bool;   // Read Product ID
      productText : Bool;   // Read Product Text
      serialNumber : Bool;   // Read Serial Number
      hwRevision : Bool;   // Read HW-Revision
      fwRevision : Bool;   // Read FW-Revision
      appSpecificName : Bool;   // Read/Write Application Specific Name
      diagnosis : Bool;   // Read diagnostics
      actualConfig : Bool;   // Read actual configuration
      targetConfig : Bool;   // Read/Write target configuration
   END_VAR
   VAR_OUTPUT
      done : Bool;   // TRUE: Commanded functionality has been completed successfully
      busy : Bool;   // TRUE: FB is not finished and new output values can be expected
      error : Bool;   // TRUE: An error occurred during the execution of the FB
      status : Word;   // 16#0000 - 16#7FFF: Status of the FB, 16#8000 - 16#FFFF: Error identification
      diagnostics : "LIOLink_typeDiagnostics";   // Diagnostics information of LIOLink_Device
   END_VAR
   VAR_IN_OUT
      data : "LIOLink_3RA_typeAll";   // Data area, device specific (Data Type)
   END_VAR
   VAR
      instDevice : "LIOLink_Device";
      statRecordParam : Struct   // Parameters to read/write specific records
         index : Array[0..#HIGHEST_REQUEST_NUMBER] of Int;   // Index of data set
         subindex : Array[0..#HIGHEST_REQUEST_NUMBER] of Int;   // Subindex of data sets
         length : Array[0..#HIGHEST_REQUEST_NUMBER] of Int;   // Length of data set
      END_STRUCT;
      statRecord : Array[0..#UPPER_BOUND_RECORD] of Byte;   // Record buffer
      statIndex : Int;   // Requested index
      statSubindex : Int;   // Requested subindex
      statRecordLen : Int;   // Length of record to be written
      statHwID : HW_IO;   // Static value for input 'hwID'
      statCap : Int;   // Static value for input 'cap'
      statReadWrite : Bool;   // Static value for input 'readWrite'
      statPort : Int;   // Static value for input 'port'
      statPollingPeriod : Time := T#100MS;   // Static value for input 'pollingPeriod'
      statParameterPage0 : Bool;   // Static value for input 'parameterPage0'
      statParameterPage1 : Bool;   // Static value for input 'parameterPage1'
      statVendorName : Bool;   // Static value for input 'vendorName'
      statVendorText : Bool;   // Static value for input 'vendorText'
      statProductName : Bool;   // Static value for input 'productName'
      statProductID : Bool;   // Static value for input 'productID'
      statProductText : Bool;   // Static value for input 'productText'
      statSerialNumber : Bool;   // Static value for input 'serialNumber'
      statHwRevision : Bool;   // Static value for input 'hwRevision'
      statFwRevision : Bool;   // Static value for input 'fwRevision'
      statAppSpecificName : Bool;   // Static value for input 'appSpecificName'
      statDiagnosis : Bool;   // Static value for input 'diagnosis'
      statActualConfig : Bool;   // Static value for input 'actualConfig'
      statTargetConfig : Bool;   // Static value for input 'targetConfig'
      statRequest : Int;   // Case of request (data set)
      statDoneOld : Bool;   // Last cycle's value of instDevice.done
   END_VAR
   VAR_TEMP
      tempIndex : Int;   // Loop index
      tempLen : UInt;   // Length
      tempRetValDeserialize : Int;   // Auxiliary tag for Deserialize RetVal
      tempRetValSerialize : Int;   // Auxiliary tag for Serialize RetVal
      tempPosDeserialize : DInt;   // Auxiliary tag for Deserialize POS Output
      tempPosSerialize : DInt;   // Auxiliary tag for Serialize POS Output
      tempFieldParameterPage0 : Array[0..#UPPER_BOUND_PARAMETER_PAGE] of Byte;   // Auxiliary tag for Parameter Page 0 record conversion
      tempFieldParameterPage1 : Array[0..#UPPER_BOUND_PARAMETER_PAGE] of Byte;   // Auxiliary tag for Parameter Page 1 record conversion
      tempFieldDiagnostics : Array[0..#UPPER_BOUND_DIAGNOSTICS] of Byte;   // Auxiliary tag for Diagnostics record conversion
      tempFieldActualConfig : Array[0..#UPPER_BOUND_ACTUAL_TARGET_CONFIG] of Byte;   // Auxiliary tag for Actual Configuration record conversion
      tempFieldTargetConfig : Array[0..#UPPER_BOUND_ACTUAL_TARGET_CONFIG] of Byte;   // Auxiliary tag for Target Configuration record conversion
      tempInternalError : Bool;   // Auxiliary tag to collect serialize and Deserialize issues
   END_VAR
   VAR CONSTANT
      UPPER_BOUND_RECORD : Int := 231;   // Upper Bound of record buffer
      HIGHEST_REQUEST_NUMBER : Int := 28;   // Highest available request number
      UPPER_BOUND_PARAMETER_PAGE : Int := 15;   // Upper Bound of Parameter Page 0 auxiliary field
      UPPER_BOUND_DIAGNOSTICS : Int := 51;   // Upper Bound of Diagnostics auxiliary field
      UPPER_BOUND_ACTUAL_TARGET_CONFIG : Int := 41;   // Upper Bound of Actual and Target Configuration auxiliary field
      MODE_READ : Bool := FALSE;   // Mode to read data
      MODE_WRITE : Bool := TRUE;   // Mode to write data
      STATUS_IDLE : Word := 16#7000;   // Status: Idle
      STATUS_EXECUTION_FINISHED : Word := 16#0000;   // Execution finished without errors
      ERR_INCONSISTENT_DATA : Word := 16#8402;   // Error: Read data record doesn't match request
      INDEX_DIRECT_PARAM0 : Int := 0;   // Record Index
      INDEX_DIRECT_PARAM1 : Int := 1;   // Record Index
      INDEX_VENDOR_NAME : Int := 16;   // Record Index
      INDEX_VENDOR_TEXT : Int := 17;   // Record Index
      INDEX_PRODUCT_NAME : Int := 18;   // Record Index
      INDEX_PRODUCT_ID : Int := 19;   // Record Index
      INDEX_PRODUCT_TEXT : Int := 20;   // Record Index
      INDEX_SERIAL_NUMBER : Int := 21;   // Record Index
      INDEX_HARDWARE_REVISION : Int := 22;   // Record Index
      INDEX_FIRMWARE_REVISION : Int := 23;   // Record Index
      INDEX_APP_SPECIFIC_NAME : Int := 24;   // Record Index
      INDEX_DIAGNOSTICS : Int := 90;   // Record Index
      INDEX_ACTUAL_CONFIG : Int := 105;   // Record Index
      INDEX_TARGET_CONFIG : Int := 130;   // Record Index
      LENGTH_DIRECT_PARAM0 : Int := 16;   // Record Length
      LENGTH_DIRECT_PARAM1 : Int := 16;   // Record Length
      LENGTH_VENDOR_NAME : Int := 10;   // Record Length
      LENGTH_VENDOR_TEXT : Int := 58;   // Record Length
      LENGTH_PRODUCT_NAME : Int := 30;   // Record Length
      LENGTH_PRODUCT_ID : Int := 8;   // Record Length
      LENGTH_PRODUCT_TEXT : Int := 2;   // Record Length
      LENGTH_SERIAL_NUMBER : Int := 8;   // Record Length
      LENGTH_HARDWARE_REVISION : Int := 4;   // Record Length
      LENGTH_FIRMWARE_REVISION : Int := 4;   // Record Length
      LENGTH_APP_SPECIFIC_NAME : Int := 32;   // Record Length
      LENGTH_DIAGNOSTICS : Int := 52;   // Record Length
      LENGTH_ACTUAL_TARGET_CONFIG : Int := 42;   // Record Length
      LENGTH_WRITE_TARGET_CONFIG : Int := 43;   // Record Length
      EMPTY_CHAR : Char := '$00';   // Default empty char to fill empty field entries
      DEVICE_TIMEOUT : Time := T#20S;   // Timeout value for the IO-Link Device Instance
   END_VAR
   // statRecordParam.index[0] := 0;
   // statRecordParam.index[1] := 0;
   // statRecordParam.index[2] := 1;
   // statRecordParam.index[3] := 0;
   // statRecordParam.index[4] := 0;
   // statRecordParam.index[5] := 0;
   // statRecordParam.index[6] := 0;
   // statRecordParam.index[7] := 0;
   // statRecordParam.index[8] := 0;
   // statRecordParam.index[9] := 0;
   // statRecordParam.index[10] := 16;
   // statRecordParam.index[11] := 17;
   // statRecordParam.index[12] := 18;
   // statRecordParam.index[13] := 19;
   // statRecordParam.index[14] := 20;
   // statRecordParam.index[15] := 21;
   // statRecordParam.index[16] := 22;
   // statRecordParam.index[17] := 23;
   // statRecordParam.index[18] := 24;
   // statRecordParam.index[19] := 0;
   // statRecordParam.index[20] := 0;
   // statRecordParam.index[21] := 0;
   // statRecordParam.index[22] := 0;
   // statRecordParam.index[23] := 90;
   // statRecordParam.index[24] := 0;
   // statRecordParam.index[25] := 0;
   // statRecordParam.index[26] := 105;
   // statRecordParam.index[27] := 130;
   // statRecordParam.index[28] := 0;
   // statRecordParam.length[0] := 0;
   // statRecordParam.length[1] := 16;
   // statRecordParam.length[2] := 16;
   // statRecordParam.length[3] := 0;
   // statRecordParam.length[4] := 0;
   // statRecordParam.length[5] := 0;
   // statRecordParam.length[6] := 0;
   // statRecordParam.length[7] := 0;
   // statRecordParam.length[8] := 0;
   // statRecordParam.length[9] := 0;
   // statRecordParam.length[10] := 10;
   // statRecordParam.length[11] := 58;
   // statRecordParam.length[12] := 30;
   // statRecordParam.length[13] := 8;
   // statRecordParam.length[14] := 2;
   // statRecordParam.length[15] := 8;
   // statRecordParam.length[16] := 4;
   // statRecordParam.length[17] := 4;
   // statRecordParam.length[18] := 32;
   // statRecordParam.length[19] := 0;
   // statRecordParam.length[20] := 0;
   // statRecordParam.length[21] := 0;
   // statRecordParam.length[22] := 0;
   // statRecordParam.length[23] := 52;
   // statRecordParam.length[24] := 0;
   // statRecordParam.length[25] := 0;
   // statRecordParam.length[26] := 42;
   // statRecordParam.length[27] := 43;
   // statRecordParam.length[28] := 0;
BEGIN
   REGION BLOCK INFO HEADER
       //===============================================================================
       // Siemens / (c)Copyright 2022
       //-------------------------------------------------------------------------------
       // Title:            LIOLink_3RA
       // Function:         Capsule block to communicate with 3RA devices
       // Library:          LIOLink
       // Author:           Siemens Industry Online Support
       // Tested with:      CPU 1513-1 PN FW 2.8
       // Engineering:      TIA Portal V16
       // Restrictions:     --
       // Requirements:     --
       //-------------------------------------------------------------------------------
       // Change log table:
       // Version  | Date       | Expert in charge       | Changes applied
       //----------|------------|------------------------|------------------------------
       // 01.00.00 | 11.04.2014 | Online Support         | First release
       // 02.00.00 | 30.03.2015 | Online Support         | Upgrade to TIA Portal V13 SP1, use function IO_LINK_DEVICE, only one function for S7-1200 and 1500
       // 02.01.00 | 23.10.2015 | Online Support         | Update to IO_LINK_DEVICE V3.1.0
       // 03.00.00 | 22.09.2020 | Online Support         | Rewrote block for FB "LIOLink_Device" V4.0.0
       // 03.01.00 | 05.10.2022 | SUP SPH                | Optimization
       //===============================================================================
   END_REGION

   REGION INIT
       IF (#execute = TRUE AND #instDevice.status = #STATUS_IDLE) THEN

           REGION Inputs
               //save inputs
               #statHwID := #hwID;
               #statCap := #cap;
               #statReadWrite := #readWrite;
               #statPort := #port;
               #statPollingPeriod := #pollingPeriod;
               #statParameterPage0 := #parameterPage0;
               #statParameterPage1 := #parameterPage1;
               #statVendorName := #vendorName;
               #statVendorText := #vendorText;
               #statProductName := #productName;
               #statProductID := #productID;
               #statProductText := #productText;
               #statSerialNumber := #serialNumber;
               #statHwRevision := #hwRevision;
               #statFwRevision := #fwRevision;
               #statAppSpecificName := #appSpecificName;
               #statDiagnosis := #diagnosis;
               #statActualConfig := #actualConfig;
               #statTargetConfig := #targetConfig;
           END_REGION

           REGION Request selector
               //set Index and RecordLen based on the request
               IF #statParameterPage0 THEN
                   #statIndex := #INDEX_DIRECT_PARAM0;
                   #statRecordLen := #LENGTH_DIRECT_PARAM0;
               ELSIF #statParameterPage1 THEN
                   #statIndex := #INDEX_DIRECT_PARAM1;
                   #statRecordLen := #LENGTH_DIRECT_PARAM1;
               ELSIF #statVendorName THEN
                   #statIndex := #INDEX_VENDOR_NAME;
                   #statRecordLen := #LENGTH_VENDOR_NAME;
               ELSIF #statVendorText THEN
                   #statIndex := #INDEX_VENDOR_TEXT;
                   #statRecordLen := #LENGTH_VENDOR_TEXT;
               ELSIF #statProductName THEN
                   #statIndex := #INDEX_PRODUCT_NAME;
                   #statRecordLen := #LENGTH_PRODUCT_NAME;
               ELSIF #statProductID THEN
                   #statIndex := #INDEX_PRODUCT_ID;
                   #statRecordLen := #LENGTH_PRODUCT_ID;
               ELSIF #statProductText THEN
                   #statIndex := #INDEX_PRODUCT_TEXT;
                   #statRecordLen := #LENGTH_PRODUCT_TEXT;
               ELSIF #statSerialNumber THEN
                   #statIndex := #INDEX_SERIAL_NUMBER;
                   #statRecordLen := #LENGTH_SERIAL_NUMBER;
               ELSIF #statHwRevision THEN
                   #statIndex := #INDEX_HARDWARE_REVISION;
                   #statRecordLen := #LENGTH_HARDWARE_REVISION;
               ELSIF #statFwRevision THEN
                   #statIndex := #INDEX_FIRMWARE_REVISION;
                   #statRecordLen := #LENGTH_FIRMWARE_REVISION;
               ELSIF #statAppSpecificName THEN
                   #statIndex := #INDEX_APP_SPECIFIC_NAME;
                   #statRecordLen := #LENGTH_APP_SPECIFIC_NAME;
               ELSIF #statDiagnosis THEN
                   #statIndex := #INDEX_DIAGNOSTICS;
                   #statRecordLen := #LENGTH_DIAGNOSTICS;  // The length in manual is a odd number (currently 53) as the last byte is empty, a even number (52) off bytes is used to have an optimized data access
               ELSIF #statActualConfig THEN
                   #statIndex := #INDEX_ACTUAL_CONFIG;
                   #statRecordLen := #LENGTH_ACTUAL_TARGET_CONFIG;
               ELSIF #statTargetConfig THEN
                   #statIndex := #INDEX_TARGET_CONFIG;
                   IF #statReadWrite = #MODE_READ THEN
                       #statRecordLen := #LENGTH_ACTUAL_TARGET_CONFIG; // It is not a fault to use the lenght of the actual config as actual and target structure are the same - for read job it is okay to use the same even length
                   ELSE
                       #statRecordLen := #LENGTH_WRITE_TARGET_CONFIG; // For write job the full data set need to be written to get accepted (currently 43 Byte) but as it is a odd structure and the last bytes are empty, internally a shorter and even structure is used 
                   END_IF;
               ELSE

                   RETURN;
               END_IF;
           END_REGION

           IF #statReadWrite = #MODE_WRITE THEN
               //prepare statRecord in case of a writing request
               REGION write
                   IF #statParameterPage1 THEN
                       #tempRetValSerialize := Serialize(SRC_VARIABLE := #data.parameterPage1, DEST_ARRAY => #tempFieldParameterPage1, POS := #tempPosSerialize);
                       UMOVE_BLK(IN := #tempFieldParameterPage1[0],
                                 COUNT := INT_TO_ULINT(#statRecordLen),
                                 OUT => #statRecord[0]);

                   ELSIF #statAppSpecificName THEN
                       Strg_TO_Chars(Strg := #data.appSpecificName,
                                     pChars := 0,
                                     Cnt => #tempLen,
                                     Chars := #statRecord);

                       // Fill remaining characters with null
                       FOR #tempIndex := UINT_TO_INT(#tempLen) TO #statRecordLen - 1 DO
                           #statRecord[#tempIndex] := CHAR_TO_BYTE(#EMPTY_CHAR);
                       END_FOR;

                   ELSIF #statTargetConfig THEN
                       // IMPORTANT: The write job and the data preparation is special as internally the data structure of the target config has a length of 42 byte for optimized handling.
                       // But the data set in the 3RA has a odd length of 43 byte.

                       #tempRetValSerialize := Serialize(SRC_VARIABLE := #data.targetConfig, DEST_ARRAY => #tempFieldTargetConfig, POS := #tempPosSerialize);
                       UMOVE_BLK(IN := #tempFieldTargetConfig[0],
                                 COUNT := INT_TO_ULINT(#LENGTH_ACTUAL_TARGET_CONFIG), // Only the netto data range (currently 42 Bytes) is copied to the record area
                                 OUT => #statRecord[0]);
                       #statRecord[#LENGTH_ACTUAL_TARGET_CONFIG] := 16#00;  // The last odd byte of the record area (Byte 43 = Index 42 in the record field) is reset to 0 as 43 Bytes need to be written as the data set is 43 Bytes long
                   ELSE // all other data sets are read only  
                       ;
                   END_IF;
                   #tempInternalError := #tempRetValSerialize <> WORD_TO_INT(#STATUS_EXECUTION_FINISHED);
               END_REGION
           END_IF;
       END_IF;
   END_REGION

   REGION CALL
       //IOL-Call -> Request to read/write from an IO-Link-Device
       #instDevice(execute := #execute,
                   hwID := #statHwID,
                   cap := #statCap,
                   readWrite := #statReadWrite,
                   "port" := #statPort,
                   pollingPeriod := #statPollingPeriod,
                   index := #statIndex,
                   subindex := #statSubindex,
                   writeLen := #statRecordLen,
                   timeout := #DEVICE_TIMEOUT,
                   record := #statRecord);
   END_REGION

   REGION READ
       // Copy data if available and valid
       IF #instDevice.done = TRUE AND #statDoneOld = FALSE AND #statReadWrite = #MODE_READ THEN
           IF #statParameterPage0 THEN
               UMOVE_BLK(IN := #statRecord[0],
                         COUNT := INT_TO_ULINT(#statRecordLen),
                         OUT => #tempFieldParameterPage0[0]);
               #tempRetValDeserialize := Deserialize(SRC_ARRAY := #tempFieldParameterPage0, DEST_VARIABLE => #data.parameterPage0, POS := #tempPosDeserialize);
           ELSIF #statParameterPage1 THEN
               UMOVE_BLK(IN := #statRecord[0],
                         COUNT := INT_TO_ULINT(#statRecordLen),
                         OUT => #tempFieldParameterPage1[0]);
               #tempRetValDeserialize := Deserialize(SRC_ARRAY := #tempFieldParameterPage1, DEST_VARIABLE => #data.parameterPage1, POS := #tempPosDeserialize);
           ELSIF #statVendorName THEN
               Chars_TO_Strg(Chars := #statRecord,
                             pChars := 0,
                             Cnt := INT_TO_UINT(#statRecordLen),
                             Strg => #data.vendorName);
           ELSIF #statVendorText THEN
               Chars_TO_Strg(Chars := #statRecord,
                             pChars := 0,
                             Cnt := INT_TO_UINT(#statRecordLen),
                             Strg => #data.vendorText);
           ELSIF #statProductName THEN
               Chars_TO_Strg(Chars := #statRecord,
                             pChars := 0,
                             Cnt := INT_TO_UINT(#statRecordLen),
                             Strg => #data.productName);
           ELSIF #statProductID THEN
               Chars_TO_Strg(Chars := #statRecord,
                             pChars := 0,
                             Cnt := INT_TO_UINT(#statRecordLen),
                             Strg => #data.productID);
           ELSIF #statProductText THEN
               Chars_TO_Strg(Chars := #statRecord,
                             pChars := 0,
                             Cnt := INT_TO_UINT(#statRecordLen),
                             Strg => #data.productText);
           ELSIF #statSerialNumber THEN
               Chars_TO_Strg(Chars := #statRecord,
                             pChars := 0,
                             Cnt := INT_TO_UINT(#statRecordLen),
                             Strg => #data.serialNumber);
           ELSIF #statHwRevision THEN
               Chars_TO_Strg(Chars := #statRecord,
                             pChars := 0,
                             Cnt := INT_TO_UINT(#statRecordLen),
                             Strg => #data.hwRevision);
           ELSIF #statFwRevision THEN
               Chars_TO_Strg(Chars := #statRecord,
                             pChars := 0,
                             Cnt := INT_TO_UINT(#statRecordLen),
                             Strg => #data.fwRevision);
           ELSIF #statAppSpecificName THEN
               Chars_TO_Strg(Chars := #statRecord,
                             pChars := 0,
                             Cnt := INT_TO_UINT(#statRecordLen),
                             Strg => #data.appSpecificName);
           ELSIF #statDiagnosis THEN
               UMOVE_BLK(IN := #statRecord[0],
                         COUNT := INT_TO_ULINT(#statRecordLen),
                         OUT => #tempFieldDiagnostics[0]);
               #tempRetValDeserialize := Deserialize(SRC_ARRAY := #tempFieldDiagnostics, DEST_VARIABLE => #data.diagnostics, POS := #tempPosDeserialize);
           ELSIF #statActualConfig THEN
               UMOVE_BLK(IN := #statRecord[0],
                         COUNT := INT_TO_ULINT(#statRecordLen),
                         OUT => #tempFieldActualConfig[0]);
               #tempRetValDeserialize := Deserialize(SRC_ARRAY := #tempFieldActualConfig, DEST_VARIABLE => #data.actualConfig, POS := #tempPosDeserialize);
           ELSIF #statTargetConfig THEN
               UMOVE_BLK(IN := #statRecord[0],
                         COUNT := INT_TO_ULINT(#statRecordLen),
                         OUT => #tempFieldTargetConfig[0]);
               #tempRetValDeserialize := Deserialize(SRC_ARRAY := #tempFieldTargetConfig, DEST_VARIABLE => #data.targetConfig, POS := #tempPosDeserialize);
           ELSE  // all other data set are not defined
               ;
           END_IF;
           #tempInternalError := #tempRetValDeserialize <> WORD_TO_INT(#STATUS_EXECUTION_FINISHED);
       END_IF;
       #statDoneOld := #instDevice.done;
   END_REGION

   REGION OUTPUTS
       IF #tempInternalError THEN //Error occured
           #done := false;
           #busy := false;
           #error := true;
           #status := #ERR_INCONSISTENT_DATA;
       ELSE //Execute successful
           #done := #instDevice.done;
           #busy := #instDevice.busy;
           #error := #instDevice.error;
           #status := #instDevice.status;
           #diagnostics := #instDevice.diagnostics;
       END_IF;
   END_REGION
END_FUNCTION_BLOCK

FUNCTION_BLOCK "LIOLink_3RB24"   // FB5110, SCL
TITLE = LIOLink_3RB24 / IO_LINK_3RB24_1500
{ S7_Optimized_Access := 'TRUE' }
AUTHOR : SIOS
FAMILY : LIOLink
VERSION : 3.1
// IO-Link Device FB for SIRIUS 3RB24  to use with S7-1200/1500 controllers! / IO-Link Geraete FB fuer SIRIUS 3RB24 zur Nutzung mit S7-1500!
   VAR_INPUT
      execute : Bool;   // Request to execute function
      cap : Int;   // Client Access Point (CAP) 0xB400 or 0x00E3 (227)
      hwID : HW_IO;   // Hardware identifier of IO-Link master module or first sub module
      readWrite : Bool;   // FALSE: read, TRUE: write
      port : Int;   // Port of the IO-Link Master for the Device
      pollingPeriod : Time := T#100MS;   // Time period of polling
      parameterPage0 : Bool;   // Read access on parameter page 0
      vendorName : Bool;   // Read vendor name
      vendorText : Bool;   // Read vendor text
      productName : Bool;   // Read product name
      productID : Bool;   // Read product ID
      productText : Bool;   // Read product text
      serialNumber : Bool;   // Read serial number
      hwRevision : Bool;   // Read hardware revision
      fwRevision : Bool;   // Read firmware revision
      appSpecificName : Bool;   // Read/Write application specific name
      processInput : Bool;   // Read input data
      processOutput : Bool;   // Read output data
      diagnosis : Bool;   // Read diagnostics
      measurements : Bool;   // Read measured values
      presetConfig : Bool;   // Read/Write preset configuration of device
      techFunctions : Bool;   // Read technology functions
   END_VAR
   VAR_OUTPUT
      done : Bool;   // TRUE: Commanded functionality has been completed successfully
      busy : Bool;   // TRUE: FB is not finished and new output values can be expected
      error : Bool;   // TRUE: An error occurred during the execution of the FB
      status : Word;   // 16#0000 - 16#7FFF: Status of the FB, 16#8000 - 16#FFFF: Error identification
      diagnostics : "LIOLink_typeDiagnostics";   // Diagnostics information of LIOLink_Device
   END_VAR
   VAR_IN_OUT
      data : "LIOLink_3RB24_typeAll";   // Data area, device specific (Data Type)
   END_VAR
   VAR
      instDevice : "LIOLink_Device";
      statRecord : Array[0..#UPPER_BOUND_RECORD] of Byte;   // Record buffer
      statIndex : Int;   // Requested index
      statSubindex : Int;   // Requested subindex
      statRecordLen : Int;   // Length of record to be written
      statHwID : HW_IO;   // Static value for input 'hwID'
      statCap : Int;   // Static value for input 'cap'
      statReadWrite : Bool;   // Static value for input 'readWrite'
      statPort : Int;   // Static value for input 'port'
      statPollingPeriod : Time := T#100MS;   // Static value for input 'pollingPeriod'
      statParameterPage0 : Bool;   // Static value for input 'parameterPage0'
      statVendorName : Bool;   // Static value for input 'vendorName'
      statVendorText : Bool;   // Static value for input 'vendorText'
      statProductName : Bool;   // Static value for input 'productName'
      statProductID : Bool;   // Static value for input 'productID'
      statProductText : Bool;   // Static value for input 'productText'
      statSerialNumber : Bool;   // Static value for input 'serialNumber'
      statHwRevision : Bool;   // Static value for input 'hwRevision'
      statFwRevision : Bool;   // Static value for input 'fwRevision'
      statAppSpecificName : Bool;   // Static value for input 'appSpecificName'
      statProcessInput : Bool;   // Static value for input 'processInput'
      statProcessOutput : Bool;   // Static value for input 'processOutput'
      statDiagnosis : Bool;   // Static value for input 'diagnosis'
      statMeasurements : Bool;   // Static value for input 'measurements'
      statPresetConfig : Bool;   // Static value for input 'presetConfig'
      statTechFunctions : Bool;   // Static value for input 'techFunctions'
      statRequest : Int;   // Case of request (data set)
      statDoneOld : Bool;   // Last cycle's value of instDevice.done
   END_VAR
   VAR_TEMP
      tempIndex : Int;   // Loop index
      tempLen : UInt;   // Record Length
      tempRetValSerialize : Int;   // Auxiliary tag for Serialize RetVal
      tempRetValDeserialize : Int;   // Auxiliary tag for Deserialize RetVal
      tempPosSerialize : DInt;   // Auxiliary tag for Serialize POS Output
      tempPosDeserialize : DInt;   // Auxiliary tag for Deserialize POS Output
      tempFieldParameterPage0 : Array[0..#UPPER_BOUND_PARAMETER_PAGE0] of Byte;   // Auxiliary tag for Parameter page 0 record conversion
      tempFieldDiagnostics : Array[0..#UPPER_BOUND_DIAGNOSTICS] of Byte;   // Auxiliary tag for Diagnostics record conversion
      tempFieldMeasuredValues : Array[0..#UPPER_BOUND_MEASURED_VALUES] of Byte;   // Auxiliary tag for Measurement record conversion
      tempFieldPresetConfig : Array[0..#UPPER_BOUND_PRESET_CONFIG] of Byte;   // Auxiliary tag for Preset record conversion
      tempFieldTechFunctions : Array[0..#UPPER_BOUND_TECH_FUNCTIONS] of Byte;   // Auxiliary tag for Technological Functions record conversion
      tempInternalError : Bool;   // Auxiliary tag to collect serialize and Deserialize issues
   END_VAR
   VAR CONSTANT
      UPPER_BOUND_RECORD : Int := 231;   // Upper Bound of record buffer
      HIGHEST_REQUEST_NUMBER : Int := 28;   // Highest available request number
      UPPER_BOUND_PARAMETER_PAGE0 : Int := 15;   // Upper Bound of Parameter Page 0 auxiliary field
      UPPER_BOUND_DIAGNOSTICS : Int := 25;   // Upper Bound of Diagnostics auxiliary field
      UPPER_BOUND_MEASURED_VALUES : Int := 39;   // Upper Bound of measured values auxiliary field
      UPPER_BOUND_PRESET_CONFIG : Int := 21;   // Upper Bound of preset configuration auxiliary field
      UPPER_BOUND_TECH_FUNCTIONS : Int := 25;   // Upper Bound of technology funtions auxiliary field
      MODE_READ : Bool := FALSE;   // Mode to read data
      MODE_WRITE : Bool := TRUE;   // Mode to write data
      STATUS_IDLE : Word := 16#7000;   // Status: Idle
      STATUS_EXECUTION_FINISHED : Word := 16#0000;   // Execution finished without errors
      ERR_INCONSISTENT_DATA : Word := 16#8402;   // Error: Read data record doesn't match request
      INDEX_DIRECT_PARAM0 : Int := 0;   // Record Index
      INDEX_VENDOR_NAME : Int := 16;   // Record Index
      INDEX_VENDOR_TEXT : Int := 17;   // Record Index
      INDEX_PRODUCT_NAME : Int := 18;   // Record Index
      INDEX_PRODUCT_ID : Int := 19;   // Record Index
      INDEX_PRODUCT_TEXT : Int := 20;   // Record Index
      INDEX_SERIAL_NUMBER : Int := 21;   // Record Index
      INDEX_HARDWARE_REVISION : Int := 22;   // Record Index
      INDEX_FIRMWARE_REVISION : Int := 23;   // Record Index
      INDEX_APP_SPECIFIC_NAME : Int := 24;   // Record Index
      INDEX_PROCESS_INPUT : Int := 40;   // Record Index
      INDEX_PROCESS_OUTPUT : Int := 41;   // Record Index
      INDEX_DIAGNOSTICS : Int := 92;   // Record Index
      INDEX_MEASUREMENTS : Int := 94;   // Record Index
      INDEX_PRESET_CONFIG : Int := 130;   // Record Index
      INDEX_TECH_FUNCTIONS : Int := 131;   // Record Index
      LENGTH_DIRECT_PARAM0 : Int := 16;   // Record Length
      LENGTH_VENDOR_NAME : Int := 10;   // Record Length
      LENGTH_VENDOR_TEXT : Int := 64;   // Record Length
      LENGTH_PRODUCT_NAME : Int := 30;   // Record Length
      LENGTH_PRODUCT_ID : Int := 12;   // Record Length
      LENGTH_PRODUCT_TEXT : Int := 2;   // Record Length
      LENGTH_SERIAL_NUMBER : Int := 8;   // Record Length
      LENGTH_HARDWARE_REVISION : Int := 4;   // Record Length
      LENGTH_FIRMWARE_REVISION : Int := 4;   // Record Length
      LENGTH_APP_SPECIFIC_NAME : Int := 32;   // Record Length
      LENGTH_PROCESS_INPUT : Int := 2;   // Record Length
      LENGTH_PROCESS_OUTPUT : Int := 1;   // Record Length
      LENGTH_DIAGNOSTICS : Int := 25;   // Record Length
      LENGTH_MEASUREMENTS : Int := 40;   // Record Length
      LENGTH_PRESET_CONFIG : Int := 22;   // Record Length
      LENGTH_TECH_FUNCTIONS : Int := 26;   // Record Length
      EMPTY_CHAR : Char := '$00';   // Default empty char to fill empty field entries
      DEVICE_TIMEOUT : Time := T#20S;   // Timeout value for the IO-Link Device Instance
   END_VAR
BEGIN
   REGION BLOCK INFO HEADER
       //===============================================================================
       // Siemens / (c)Copyright 2022
       //-------------------------------------------------------------------------------
       // Title:            LIOLink_3RB24
       // Function:         Capsule block to communicate with 3RB24 devices
       // Library:          LIOLink
       // Author:           Siemens Industry Online Support
       // Tested with:      CPU 1513-1 PN FW 2.8
       // Engineering:      TIA Portal V16
       // Restrictions:     --
       // Requirements:     --
       //-------------------------------------------------------------------------------
       // Change log table:
       // Version  | Date       | Expert in charge       | Changes applied
       //----------|------------|------------------------|------------------------------
       // 01.00.00 | 11.04.2014 | Online Support         | First release
       // 02.00.00 | 30.03.2015 | Online Support         | Upgrade to TIA Portal V13 SP1, use function IO_LINK_DEVICE, only one function for S7-1200 and 1500
       // 02.01.00 | 23.10.2015 | Online Support         | Update to IO_LINK_DEVICE Version 3.1
       // 03.00.00 | 01.09.2020 | Online Support         | Upgraded FB "LIOLink_Device" to V4.0.0
       // 03.01.00 | 05.10.2022 | SUP SPH                | Optimization   
       //===============================================================================
   END_REGION

   REGION INIT
       IF (#execute = TRUE AND #instDevice.status = #STATUS_IDLE) THEN

           REGION Inputs
               //save inputs
               #statHwID := #hwID;
               #statCap := #cap;
               #statReadWrite := #readWrite;
               #statPort := #port;
               #statPollingPeriod := #pollingPeriod;
               #statParameterPage0 := #parameterPage0;
               #statVendorName := #vendorName;
               #statVendorText := #vendorText;
               #statProductName := #productName;
               #statProductID := #productID;
               #statProductText := #productText;
               #statSerialNumber := #serialNumber;
               #statHwRevision := #hwRevision;
               #statFwRevision := #fwRevision;
               #statAppSpecificName := #appSpecificName;
               #statProcessInput := #processInput;
               #statProcessOutput := #processOutput;
               #statDiagnosis := #diagnosis;
               #statMeasurements := #measurements;
               #statPresetConfig := #presetConfig;
               #statTechFunctions := #techFunctions;
           END_REGION

           REGION Request selector
               //set Index and RecordLen based on the request
               IF #statParameterPage0 THEN
                   #statIndex := #INDEX_DIRECT_PARAM0;
                   #statRecordLen := #LENGTH_DIRECT_PARAM0;
               ELSIF #statVendorName THEN
                   #statIndex := #INDEX_VENDOR_NAME;
                   #statRecordLen := #LENGTH_VENDOR_NAME;
               ELSIF #statVendorText THEN
                   #statIndex := #INDEX_VENDOR_TEXT;
                   #statRecordLen := #LENGTH_VENDOR_TEXT;
               ELSIF #statProductName THEN
                   #statIndex := #INDEX_PRODUCT_NAME;
                   #statRecordLen := #LENGTH_PRODUCT_NAME;
               ELSIF #statProductID THEN
                   #statIndex := #INDEX_PRODUCT_ID;
                   #statRecordLen := #LENGTH_PRODUCT_ID;
               ELSIF #statProductText THEN
                   #statIndex := #INDEX_PRODUCT_TEXT;
                   #statRecordLen := #LENGTH_PRODUCT_TEXT;
               ELSIF #statSerialNumber THEN
                   #statIndex := #INDEX_SERIAL_NUMBER;
                   #statRecordLen := #LENGTH_SERIAL_NUMBER;
               ELSIF #statHwRevision THEN
                   #statIndex := #INDEX_HARDWARE_REVISION;
                   #statRecordLen := #LENGTH_HARDWARE_REVISION;
               ELSIF #statFwRevision THEN
                   #statIndex := #INDEX_FIRMWARE_REVISION;
                   #statRecordLen := #LENGTH_FIRMWARE_REVISION;
               ELSIF #statAppSpecificName THEN
                   #statIndex := #INDEX_APP_SPECIFIC_NAME;
                   #statRecordLen := #LENGTH_APP_SPECIFIC_NAME;
               ELSIF #statProcessInput THEN
                   #statIndex := #INDEX_PROCESS_INPUT;
                   #statRecordLen := #LENGTH_PROCESS_INPUT;
               ELSIF #statProcessOutput THEN
                   #statIndex := #INDEX_PROCESS_OUTPUT;
                   #statRecordLen := #LENGTH_PROCESS_OUTPUT;
               ELSIF #statDiagnosis THEN
                   #statIndex := #INDEX_DIAGNOSTICS;
                   #statRecordLen := #LENGTH_DIAGNOSTICS;
               ELSIF #statMeasurements THEN
                   #statIndex := #INDEX_MEASUREMENTS;
                   #statRecordLen := #LENGTH_MEASUREMENTS;
               ELSIF #statPresetConfig THEN
                   #statIndex := #INDEX_PRESET_CONFIG;
                   #statRecordLen := #LENGTH_PRESET_CONFIG;
               ELSIF #statTechFunctions THEN
                   #statIndex := #INDEX_TECH_FUNCTIONS;
                   #statRecordLen := #LENGTH_TECH_FUNCTIONS;
               ELSE
                   RETURN;
               END_IF;
           END_REGION

           IF #statReadWrite = #MODE_WRITE THEN
               //prepare statRecord in case of a writing request
               REGION write
                   IF #statAppSpecificName THEN
                       Strg_TO_Chars(Strg := #data.appSpecificName,
                                     pChars := 0,
                                     Cnt => #tempLen,
                                     Chars := #statRecord);

                       // Fill remaining characters with null
                       FOR #tempIndex := UINT_TO_INT(#tempLen) TO #statRecordLen - 1 DO
                           #statRecord[#tempIndex] := CHAR_TO_BYTE(#EMPTY_CHAR);
                       END_FOR;

                   ELSIF #statPresetConfig THEN
                       #tempRetValSerialize := Serialize(SRC_VARIABLE := #data.presetConfig, DEST_ARRAY => #tempFieldPresetConfig, POS := #tempPosSerialize);
                       UMOVE_BLK(IN := #tempFieldPresetConfig[0],
                                 COUNT := INT_TO_ULINT(#statRecordLen),
                                 OUT => #statRecord[0]);
                   ELSE // all other data sets are read only  
                       ;
                   END_IF;
                   #tempInternalError := #tempRetValSerialize <> WORD_TO_INT(#STATUS_EXECUTION_FINISHED);
               END_REGION

           END_IF;
       END_IF;
   END_REGION

   REGION CALL
       //IOL-Call -> Request to read/write from an IO-Link-Device
       #instDevice(execute := #execute,
                   hwID := #statHwID,
                   cap := #statCap,
                   readWrite := #statReadWrite,
                   "port" := #statPort,
                   pollingPeriod := #statPollingPeriod,
                   index := #statIndex,
                   subindex := #statSubindex,
                   writeLen := #statRecordLen,
                   timeout := #DEVICE_TIMEOUT,
                   record := #statRecord);
   END_REGION

   REGION READ
       // Copy data if available and valid
       IF #instDevice.done = TRUE AND #statDoneOld = FALSE AND #statReadWrite = #MODE_READ THEN
           IF #statParameterPage0 THEN
               UMOVE_BLK(IN := #statRecord[0],
                         COUNT := INT_TO_ULINT(#statRecordLen),
                         OUT => #tempFieldParameterPage0[0]);
               #tempRetValDeserialize := Deserialize(SRC_ARRAY := #tempFieldParameterPage0, DEST_VARIABLE => #data.parameterPage0, POS := #tempPosDeserialize);

           ELSIF #statVendorName THEN
               Chars_TO_Strg(Chars := #statRecord,
                             pChars := 0,
                             Cnt := INT_TO_UINT(#statRecordLen),
                             Strg => #data.vendorName);

           ELSIF #statVendorText THEN
               Chars_TO_Strg(Chars := #statRecord,
                             pChars := 0,
                             Cnt := INT_TO_UINT(#statRecordLen),
                             Strg => #data.vendorText);

           ELSIF #statProductName THEN
               Chars_TO_Strg(Chars := #statRecord,
                             pChars := 0,
                             Cnt := INT_TO_UINT(#statRecordLen),
                             Strg => #data.productName);

           ELSIF #statProductID THEN
               Chars_TO_Strg(Chars := #statRecord,
                             pChars := 0,
                             Cnt := INT_TO_UINT(#statRecordLen),
                             Strg => #data.productID);

           ELSIF #statProductText THEN
               Chars_TO_Strg(Chars := #statRecord,
                             pChars := 0,
                             Cnt := INT_TO_UINT(#statRecordLen),
                             Strg => #data.productText);
           ELSIF #statSerialNumber THEN
               Chars_TO_Strg(Chars := #statRecord,
                             pChars := 0,
                             Cnt := INT_TO_UINT(#statRecordLen),
                             Strg => #data.serialNumber);

           ELSIF #statHwRevision THEN
               Chars_TO_Strg(Chars := #statRecord,
                             pChars := 0,
                             Cnt := INT_TO_UINT(#statRecordLen),
                             Strg => #data.hwRevision);
           ELSIF #statFwRevision THEN
               Chars_TO_Strg(Chars := #statRecord,
                             pChars := 0,
                             Cnt := INT_TO_UINT(#statRecordLen),
                             Strg => #data.fwRevision);

           ELSIF #statAppSpecificName THEN
               Chars_TO_Strg(Chars := #statRecord,
                             pChars := 0,
                             Cnt := INT_TO_UINT(#statRecordLen),
                             Strg => #data.appSpecificName);

           ELSIF #statProcessInput THEN
               #data.processInput.%B0 := #statRecord[0];
               #data.processInput.%B1 := #statRecord[1];

           ELSIF #statProcessOutput THEN
               #data.processOutput := #statRecord[0];

           ELSIF #statDiagnosis THEN
               UMOVE_BLK(IN := #statRecord[0],
                         COUNT := INT_TO_ULINT(#statRecordLen),
                         OUT => #tempFieldDiagnostics[0]);
               #tempRetValDeserialize := Deserialize(SRC_ARRAY := #tempFieldDiagnostics, DEST_VARIABLE => #data.diagnostics, POS := #tempPosDeserialize);

           ELSIF #statMeasurements THEN
               UMOVE_BLK(IN := #statRecord[0],
                         COUNT := INT_TO_ULINT(#statRecordLen),
                         OUT => #tempFieldMeasuredValues[0]);
               #tempRetValDeserialize := Deserialize(SRC_ARRAY := #tempFieldMeasuredValues, DEST_VARIABLE => #data.measuredValues, POS := #tempPosDeserialize);

           ELSIF #statPresetConfig THEN
               UMOVE_BLK(IN := #statRecord[0],
                         COUNT := INT_TO_ULINT(#statRecordLen),
                         OUT => #tempFieldPresetConfig[0]);
               #tempRetValDeserialize := Deserialize(SRC_ARRAY := #tempFieldPresetConfig, DEST_VARIABLE => #data.presetConfig, POS := #tempPosDeserialize);

           ELSIF #statTechFunctions THEN
               UMOVE_BLK(IN := #statRecord[0],
                         COUNT := INT_TO_ULINT(#statRecordLen),
                         OUT => #tempFieldTechFunctions[0]);
               #tempRetValDeserialize := Deserialize(SRC_ARRAY := #tempFieldTechFunctions, DEST_VARIABLE => #data.techFunctions, POS := #tempPosDeserialize);
           ELSE  // Other data sets are not defined
               ;
           END_IF;
           #tempInternalError := #tempRetValDeserialize <> WORD_TO_INT(#STATUS_EXECUTION_FINISHED);
       END_IF;

       #statDoneOld := #instDevice.done;
   END_REGION

   REGION OUTPUTS
       IF #tempInternalError THEN //Error occured
           #done := false;
           #busy := false;
           #error := true;
           #status := #ERR_INCONSISTENT_DATA;
       ELSE //Execute successful
           #done := #instDevice.done;
           #busy := #instDevice.busy;
           #error := #instDevice.error;
           #status := #instDevice.status;
           #diagnostics := #instDevice.diagnostics;
       END_IF;
   END_REGION
END_FUNCTION_BLOCK

